Fanuc KAREL source: kt00300.KL

-- PROVISIONAL review KL for V770-1; original PC SHA256 5afca9adfa75683988d3fdf210c5727fbcef32caf12140b37318d02423ab01fc
-- Incomplete behavior may be omitted. Consult companion uncertainty JSON. Do not deploy.
PROGRAM KT00300
%NOLOCKGROUP
VAR
  R1 : REAL
  OUT : BOOLEAN
-- UNRESOLVED_DECL H2 type=002017
BEGIN
  -- UNRESOLVED_PC offsets 5-16; opcodes 2E,23
  -- UNRESOLVED_PC offsets 21-35; opcodes 2E,22,9D,33,B4
  -- UNRESOLVED_PC offsets 40-63; opcodes 21,22,9D,33,B3,64,6E,23
  -- UNRESOLVED_PC offsets 68-72; opcodes 7F
END KT00300
